                                               //Partner information is already known in the diagnostic structure
                                               IF (#diagnostics.partnerConfig.connnection.lifeSignCycleTime = T#0ms) THEN
                                                   //No --> Get diagnostics information
                                                   //LCom V2
                                                   IF (#statActualLocalLComVersion = #HEADER_V2) THEN
                                                       //UsesTimeStamp
                                                       #diagnostics.partnerConfig.timeSync.usePartnerTimestamps := BYTE_TO_BOOL(#statReceive.tempTelegram.data[2]);
                                                       //SendModeSyncTime
                                                       #diagnostics.partnerConfig.timeSync.sendMode := #statReceive.tempTelegram.data[3];
                                                       //LifeSignCycle
                                                       #tempDWord.%B3 := #statReceive.tempTelegram.data[4];
                                                       #tempDWord.%B2 := #statReceive.tempTelegram.data[5];
                                                       #tempDWord.%B1 := #statReceive.tempTelegram.data[6];
                                                       #tempDWord.%B0 := #statReceive.tempTelegram.data[7];
                                                       #statReceive.configTelegramV2.lifeSignCycle := DWORD_TO_TIME(#tempDWord);
                                                       #diagnostics.partnerConfig.connnection.lifeSignCycleTime := #statReceive.configTelegramV2.lifeSignCycle;
                                                       //Sender cycleTime
                                                       #tempDWord.%B3 := #statReceive.tempTelegram.data[8];
                                                       #tempDWord.%B2 := #statReceive.tempTelegram.data[9];
                                                       #tempDWord.%B1 := #statReceive.tempTelegram.data[10];
                                                       #tempDWord.%B0 := #statReceive.tempTelegram.data[11];
                                                       #statReceive.configTelegramV2.cycleTime := DWORD_TO_TIME(#tempDWord);
                                                       #diagnostics.partnerConfig.sender.cycleTime := #statReceive.configTelegramV2.cycleTime;
                                                       //Sender ackTimeOut
                                                       #tempDWord.%B3 := #statReceive.tempTelegram.data[12];
                                                       #tempDWord.%B2 := #statReceive.tempTelegram.data[13];
                                                       #tempDWord.%B1 := #statReceive.tempTelegram.data[14];
                                                       #tempDWord.%B0 := #statReceive.tempTelegram.data[15];
                                                       #statReceive.configTelegramV2.ackTimeOut := DWORD_TO_TIME(#tempDWord);
                                                       #diagnostics.partnerConfig.sender.ackTimeout := #statReceive.configTelegramV2.ackTimeOut;
                                                       //MaxSendDataLength
                                                       #tempDWord.%B3 := #statReceive.tempTelegram.data[16];
                                                       #tempDWord.%B2 := #statReceive.tempTelegram.data[17];
                                                       #tempDWord.%B1 := #statReceive.tempTelegram.data[18];
                                                       #tempDWord.%B0 := #statReceive.tempTelegram.data[19];
                                                       #statReceive.configTelegramV2.maxSendDataLength := #tempDWord;
                                                       #diagnostics.partnerConfig.sizeOfSendBuffer := #statReceive.configTelegramV2.maxSendDataLength;
                                                       //MaxReceiveDataLength
                                                       #tempDWord.%B3 := #statReceive.tempTelegram.data[20];
                                                       #tempDWord.%B2 := #statReceive.tempTelegram.data[21];
                                                       #tempDWord.%B1 := #statReceive.tempTelegram.data[22];
                                                       #tempDWord.%B0 := #statReceive.tempTelegram.data[23];
                                                       #statReceive.configTelegramV2.maxReceiveDataLength := #tempDWord;
                                                       #diagnostics.partnerConfig.sizeOfReceiveBuffer := #statReceive.configTelegramV2.maxReceiveDataLength;
                                                   ELSE
                                                       //LCom V1
                                                       //LifeSignCycle
                                                       #statReceive.configTelegramV1.lifeSignCycle.%B1 := #statReceive.tempTelegram.data[8];
                                                       #statReceive.configTelegramV1.lifeSignCycle.%B0 := #statReceive.tempTelegram.data[9];
                                                       #diagnostics.partnerConfig.connnection.lifeSignCycleTime := UINT_TO_TIME(#statReceive.configTelegramV1.lifeSignCycle);
                                                       //MaxSendDataLength
                                                       #statReceive.configTelegramV1.maxSendDataLength.%B1 := #statReceive.tempTelegram.data[12];
                                                       #statReceive.configTelegramV1.maxSendDataLength.%B0 := #statReceive.tempTelegram.data[13];
                                                       #diagnostics.partnerConfig.sizeOfSendBuffer := #statReceive.configTelegramV1.maxSendDataLength;
                                                       //MaxReceiveDataLength
                                                       #statReceive.configTelegramV1.maxReceiveDataLength.%B1 := #statReceive.tempTelegram.data[14];
                                                       #statReceive.configTelegramV1.maxReceiveDataLength.%B0 := #statReceive.tempTelegram.data[15];
                                                       #diagnostics.partnerConfig.sizeOfReceiveBuffer := #statReceive.configTelegramV1.maxReceiveDataLength;
                                                       //UsesTimeStamp
                                                       #diagnostics.partnerConfig.timeSync.usePartnerTimestamps := BYTE_TO_BOOL(#statReceive.tempTelegram.data[10]);
                                                       //SendModeSyncTime
                                                       #diagnostics.partnerConfig.timeSync.sendMode := #statReceive.tempTelegram.data[11];
                                                   END_IF;
                                               END_IF;

                                           1://Telegram type 1

                                               //Reset index, so a new temp. LCom header can be built
                                               #statReceive.tempTelegram.index := 0;
                                               #statReceive.numberOfLComHeader := #statReceive.numberOfLComHeader + 1;

                                               //LCom V1
                                               //LifeSignCycle
                                               #statReceive.configTelegramV1.lifeSignCycle.%B1 := #statReceive.tempTelegram.data[8];
                                               #statReceive.configTelegramV1.lifeSignCycle.%B0 := #statReceive.tempTelegram.data[9];
                                               #diagnostics.partnerConfig.connnection.lifeSignCycleTime := UINT_TO_TIME(#statReceive.configTelegramV1.lifeSignCycle);
                                               //Receiver cycleTime from receiver
                                               #statReceive.configTelegramV1.cycleTime.%B1 := #statReceive.tempTelegram.data[4];
                                               #statReceive.configTelegramV1.cycleTime.%B0 := #statReceive.tempTelegram.data[5];
                                               //Receiver ackTimeOut from receiver
                                               #statReceive.configTelegramV1.ackTimeOut.%B1 := #statReceive.tempTelegram.data[6];
                                               #statReceive.configTelegramV1.ackTimeOut.%B0 := #statReceive.tempTelegram.data[7];

                                               //Are receive cycle time and current sender cycle time and receive ackTimeOut and current sender ackTimeOut equal ?
                                               IF ((#statReceive.configTelegramV1.cycleTime = (TIME_TO_UINT(#diagnostics.localConfig.sender.cycleTime)))
                                                   AND
                                                   (#statReceive.configTelegramV1.ackTimeOut = (TIME_TO_UINT(#diagnostics.localConfig.sender.ackTimeout))))
                                               THEN
                                                   ;//Yes equal --> Set FB.#connected and diagnostics information
                                               ELSE
                                                   //Not equal --> Compare values and prioritize
                                                   //Compare cycle time
                                                   IF (#statReceive.configTelegramV1.cycleTime > (TIME_TO_UINT(#diagnostics.localConfig.sender.cycleTime))) THEN
                                                       #statSend.configTelegramV1.cycleTime := #statReceive.configTelegramV1.cycleTime;
                                                   ELSE
                                                       ;//Actual sender cycleTime is bigger than the received sender cycleTime
                                                   END_IF;

                                                   //Compare acknowledge timeout
                                                   IF (#statReceive.configTelegramV1.ackTimeOut > (TIME_TO_UINT(#diagnostics.localConfig.sender.ackTimeout))) THEN
                                                       #statSend.configTelegramV1.ackTimeOut := #statReceive.configTelegramV1.ackTimeOut;
                                                   ELSE
                                                       ;//Actual acknowledge timeout is bigger than the received sender acknowledge timeout
                                                   END_IF;

                                                   //Update diagnostics information
                                                   #diagnostics.localConfig.sender.cycleTime := UINT_TO_TIME(#statReceive.configTelegramV1.cycleTime);
                                                   #diagnostics.localConfig.sender.ackTimeout := UINT_TO_TIME(#statReceive.configTelegramV1.ackTimeOut);

                                                   //Send telegram 2
                                                   #statSend.tsendFct.data[#statSend.tsendFct.dataOffset] := #statSend.configTelegramV1.LComVersion;
                                                   #statSend.tsendFct.data[#statSend.tsendFct.dataOffset + 1] := 16#02;
                                                   #statSend.tsendFct.data[#statSend.tsendFct.dataOffset + 2] := #statSend.configTelegramV1.comMode;
                                                   #statSend.tsendFct.data[#statSend.tsendFct.dataOffset + 3] := #statSend.configTelegramV1.slidingWindow;
                                                   //Cycle time
                                                   #statSend.tsendFct.data[#statSend.tsendFct.dataOffset + 4] := #statSend.configTelegramV1.cycleTime.%B1;
                                                   #statSend.tsendFct.data[#statSend.tsendFct.dataOffset + 5] := #statSend.configTelegramV1.cycleTime.%B0;
                                                   //Acknowledge timeout
                                                   #statSend.tsendFct.data[#statSend.tsendFct.dataOffset + 6] := #statSend.configTelegramV1.ackTimeOut.%B1;
                                                   #statSend.tsendFct.data[#statSend.tsendFct.dataOffset + 7] := #statSend.configTelegramV1.ackTimeOut.%B0;
                                                   //LifeSignCycle
                                                   #statSend.tsendFct.data[#statSend.tsendFct.dataOffset + 8] := #statSend.configTelegramV1.lifeSignCycle.%B1;
                                                   #statSend.tsendFct.data[#statSend.tsendFct.dataOffset + 9] := #statSend.configTelegramV1.lifeSignCycle.%B0;
                                                   //Status
                                                   #statSend.tsendFct.data[#statSend.tsendFct.dataOffset + 10] := #statSend.configTelegramV1.status;
                                                   //SendModeSyncTime
                                                   #statSend.tsendFct.data[#statSend.tsendFct.dataOffset + 11] := #statSend.configTelegramV1.sendModeSyncTime;
                                                   //MaxSendDataLength
                                                   #statSend.tsendFct.data[#statSend.tsendFct.dataOffset + 12] := #statSend.configTelegramV1.maxSendDataLength.%B1;
                                                   #statSend.tsendFct.data[#statSend.tsendFct.dataOffset + 13] := #statSend.configTelegramV1.maxSendDataLength.%B0;
                                                   //MaxReceiveDataLength
                                                   #statSend.tsendFct.data[#statSend.tsendFct.dataOffset + 14] := #statSend.configTelegramV1.maxReceiveDataLength.%B1;
                                                   #statSend.tsendFct.data[#statSend.tsendFct.dataOffset + 15] := #statSend.configTelegramV1.maxReceiveDataLength.%B0;
                                                   //Calculate offset in the tcp send buffer
                                                   #statSend.tsendFct.dataOffset := #statSend.tsendFct.dataOffset + 16;
                                                   #statState.sender := #SEND_CONFIG;
                                               END_IF;

                                               //Set FB.#connected and #diagnostics information
                                               #connected := #statConnected := TRUE;
                                               #diagnostics.statistics.LComProtocolUsed := TRUE;
                                               #diagnostics.statistics.activeLComVersion := #HEADER_V1;
                                               //Write diagnostics
                                               #statDiag.bufferIndex := #statDiag.bufferIndex + 1;
                                               #statDiag.buffer[#statDiag.bufferIndex].status := #STATUS_CONNECTED_V1;
                                               #statDiag.buffer[#statDiag.bufferIndex].subFunctionErrorID := 16#0000;
                                               #statDiag.buffer[#statDiag.bufferIndex].additionalValue1 := 0.0;
                                               #statDiag.buffer[#statDiag.bufferIndex].additionalValue2 := 0.0;
                                               #statDiag.buffer[#statDiag.bufferIndex].additionalValue3 := 0.0;
                                               #statDiag.buffer[#statDiag.bufferIndex].additionalValue4 := T#0ms;

                                               #statState.cfgSender := #OPERATION;

                                               //MaxSendDataLength
                                               #statReceive.configTelegramV1.maxSendDataLength.%B1 := #statReceive.tempTelegram.data[12];
                                               #statReceive.configTelegramV1.maxSendDataLength.%B0 := #statReceive.tempTelegram.data[13];
                                               #diagnostics.partnerConfig.sizeOfSendBuffer := #statReceive.configTelegramV1.maxSendDataLength;
                                               //MaxReceiveDataLength
                                               #statReceive.configTelegramV1.maxReceiveDataLength.%B1 := #statReceive.tempTelegram.data[14];
                                               #statReceive.configTelegramV1.maxReceiveDataLength.%B0 := #statReceive.tempTelegram.data[15];
                                               #diagnostics.partnerConfig.sizeOfReceiveBuffer := #statReceive.configTelegramV1.maxReceiveDataLength;
                                               //UsesTimeStamp
                                               #diagnostics.partnerConfig.timeSync.usePartnerTimestamps := BYTE_TO_BOOL(#statReceive.tempTelegram.data[10]);
                                               //SendModeSyncTime
                                               #diagnostics.partnerConfig.timeSync.sendMode := #statReceive.tempTelegram.data[11];

                                               IF ((#diagnostics.localConfig.timeSync.usePartnerTimestamps
                                                   XOR
                                                   #diagnostics.partnerConfig.timeSync.usePartnerTimestamps)
                                                   AND
                                                   (#diagnostics.localConfig.timeSync.sendMode > 0
                                                   OR
                                                   #diagnostics.partnerConfig.timeSync.sendMode > 0))
                                               THEN
                                                   ;//One cpu does send timeSync information
                                               ELSE
                                                   //Write diagnostics
                                                   #statDiag.bufferIndex := #statDiag.bufferIndex + 1;
                                                   #statDiag.buffer[#statDiag.bufferIndex].status := #WARN_NO_TIME_SYNC;
                                                   #statDiag.buffer[#statDiag.bufferIndex].subFunctionErrorID := 16#0000;
                                                   #statDiag.buffer[#statDiag.bufferIndex].additionalValue1 := 0.0;
                                                   #statDiag.buffer[#statDiag.bufferIndex].additionalValue2 := 0.0;
                                                   #statDiag.buffer[#statDiag.bufferIndex].additionalValue3 := 0.0;
                                                   #statDiag.buffer[#statDiag.bufferIndex].additionalValue4 := T#0ms;
                                               END_IF;

                                           2://telegram type 2

                                               //Reset index, so a new temp. LCom header can be built
                                               #statReceive.tempTelegram.index := 0;
                                               #statReceive.numberOfLComHeader := #statReceive.numberOfLComHeader + 1;

                                               //LCom V2
                                               IF (#statActualLocalLComVersion = #HEADER_V2) THEN
                                                   //UsesTimeStamp
                                                   #diagnostics.partnerConfig.timeSync.usePartnerTimestamps := BYTE_TO_BOOL(#statReceive.tempTelegram.data[2]);
                                                   //SendModeSyncTime
                                                   #diagnostics.partnerConfig.timeSync.sendMode := #statReceive.tempTelegram.data[3];
                                                   //LifeSignCycle
                                                   #tempDWord.%B3 := #statReceive.tempTelegram.data[4];
                                                   #tempDWord.%B2 := #statReceive.tempTelegram.data[5];
                                                   #tempDWord.%B1 := #statReceive.tempTelegram.data[6];
                                                   #tempDWord.%B0 := #statReceive.tempTelegram.data[7];
                                                   #statReceive.configTelegramV2.lifeSignCycle := DWORD_TO_TIME(#tempDWord);
                                                   #diagnostics.partnerConfig.connnection.lifeSignCycleTime := #statReceive.configTelegramV2.lifeSignCycle;

                                                   //Sender cycleTime
                                                   #tempDWord.%B3 := #statReceive.tempTelegram.data[8];
                                                   #tempDWord.%B2 := #statReceive.tempTelegram.data[9];
                                                   #tempDWord.%B1 := #statReceive.tempTelegram.data[10];
                                                   #tempDWord.%B0 := #statReceive.tempTelegram.data[11];
                                                   #statReceive.configTelegramV2.cycleTime := DWORD_TO_TIME(#tempDWord);
                                                   #diagnostics.partnerConfig.sender.cycleTime := #statReceive.configTelegramV2.cycleTime;
                                                   //Sender ackTimeOut
                                                   #tempDWord.%B3 := #statReceive.tempTelegram.data[12];
                                                   #tempDWord.%B2 := #statReceive.tempTelegram.data[13];
                                                   #tempDWord.%B1 := #statReceive.tempTelegram.data[14];
                                                   #tempDWord.%B0 := #statReceive.tempTelegram.data[15];
                                                   #statReceive.configTelegramV2.ackTimeOut := DWORD_TO_TIME(#tempDWord);
                                                   #diagnostics.partnerConfig.sender.ackTimeout := #statReceive.configTelegramV2.ackTimeOut;
                                                   //MaxSendDataLength
                                                   #tempDWord.%B3 := #statReceive.tempTelegram.data[16];
                                                   #tempDWord.%B2 := #statReceive.tempTelegram.data[17];
                                                   #tempDWord.%B1 := #statReceive.tempTelegram.data[18];
                                                   #tempDWord.%B0 := #statReceive.tempTelegram.data[19];
                                                   #statReceive.configTelegramV2.maxSendDataLength := #tempDWord;
                                                   #diagnostics.partnerConfig.sizeOfSendBuffer := #statReceive.configTelegramV2.maxSendDataLength;
                                                   //MaxReceiveDataLength
                                                   #tempDWord.%B3 := #statReceive.tempTelegram.data[20];
                                                   #tempDWord.%B2 := #statReceive.tempTelegram.data[21];
                                                   #tempDWord.%B1 := #statReceive.tempTelegram.data[22];
                                                   #tempDWord.%B0 := #statReceive.tempTelegram.data[23];
                                                   #statReceive.configTelegramV2.maxReceiveDataLength := #tempDWord;
                                                   #diagnostics.partnerConfig.sizeOfReceiveBuffer := #statReceive.configTelegramV2.maxReceiveDataLength;

                                                   //Set FB.#connected and #diagnostics information
                                                   #connected := #statConnected := TRUE;
                                                   #diagnostics.statistics.LComProtocolUsed := TRUE;
                                                   #diagnostics.statistics.activeLComVersion := #HEADER_V2;
                                                   #statState.cfgSender := #OPERATION;

                                                   //Write diagnostics
                                                   #statDiag.bufferIndex := #statDiag.bufferIndex + 1;
                                                   #statDiag.buffer[#statDiag.bufferIndex].status := #STATUS_CONNECTED_V2;
                                                   #statDiag.buffer[#statDiag.bufferIndex].subFunctionErrorID := 16#0000;
                                                   #statDiag.buffer[#statDiag.bufferIndex].additionalValue1 := 0.0;
                                                   #statDiag.buffer[#statDiag.bufferIndex].additionalValue2 := 0.0;
                                                   #statDiag.buffer[#statDiag.bufferIndex].additionalValue3 := 0.0;
                                                   #statDiag.buffer[#statDiag.bufferIndex].additionalValue4 := T#0ms;

                                                   //Check timeSync setting at local cpu and partner cpu
                                                   IF ((#diagnostics.localConfig.timeSync.usePartnerTimestamps
                                                       XOR
                                                       #diagnostics.partnerConfig.timeSync.usePartnerTimestamps)
                                                       AND
                                                       (#diagnostics.localConfig.timeSync.sendMode > 0
                                                       OR
                                                       #diagnostics.partnerConfig.timeSync.sendMode > 0))
                                                   THEN
                                                       ;//One cpu does send timeSync information
                                                   ELSE
                                                       //Write diagnostics
                                                       #statDiag.bufferIndex := #statDiag.bufferIndex + 1;
                                                       #statDiag.buffer[#statDiag.bufferIndex].status := #WARN_NO_TIME_SYNC;
                                                       #statDiag.buffer[#statDiag.bufferIndex].subFunctionErrorID := 16#0000;
                                                       #statDiag.buffer[#statDiag.bufferIndex].additionalValue1 := 0.0;
                                                       #statDiag.buffer[#statDiag.bufferIndex].additionalValue2 := 0.0;
                                                       #statDiag.buffer[#statDiag.bufferIndex].additionalValue3 := 0.0;
                                                       #statDiag.buffer[#statDiag.bufferIndex].additionalValue4 := T#0ms;
                                                   END_IF;
                                                   //Do not send telegram 1
                                               ELSE
                                                   //LCom V1
                                                   //LifeSignCycle
                                                   #statReceive.configTelegramV1.lifeSignCycle.%B1 := #statReceive.tempTelegram.data[8];
                                                   #statReceive.configTelegramV1.lifeSignCycle.%B0 := #statReceive.tempTelegram.data[9];
                                                   #diagnostics.partnerConfig.connnection.lifeSignCycleTime := UINT_TO_TIME(#statReceive.configTelegramV1.lifeSignCycle);
                                                   //CycleTime
                                                   #statReceive.configTelegramV1.cycleTime.%B1 := #statReceive.tempTelegram.data[4];
                                                   #statReceive.configTelegramV1.cycleTime.%B0 := #statReceive.tempTelegram.data[5];
                                                   #diagnostics.partnerConfig.sender.cycleTime := UINT_TO_TIME(#statReceive.configTelegramV1.cycleTime);
                                                   //AckTimeOut
                                                   #statReceive.configTelegramV1.ackTimeOut.%B1 := #statReceive.tempTelegram.data[6];
                                                   #statReceive.configTelegramV1.ackTimeOut.%B0 := #statReceive.tempTelegram.data[7];
                                                   #diagnostics.partnerConfig.sender.ackTimeout := UINT_TO_TIME(#statReceive.configTelegramV1.ackTimeOut);
                                                   //MaxSendDataLength
                                                   #statReceive.configTelegramV1.maxSendDataLength.%B1 := #statReceive.tempTelegram.data[12];
                                                   #statReceive.configTelegramV1.maxSendDataLength.%B0 := #statReceive.tempTelegram.data[13];
                                                   #diagnostics.partnerConfig.sizeOfSendBuffer := #statReceive.configTelegramV1.maxSendDataLength;
                                                   //MaxReceiveDataLength
                                                   #statReceive.configTelegramV1.maxReceiveDataLength.%B1 := #statReceive.tempTelegram.data[14];
                                                   #statReceive.configTelegramV1.maxReceiveDataLength.%B0 := #statReceive.tempTelegram.data[15];
                                                   #diagnostics.partnerConfig.sizeOfReceiveBuffer := #statReceive.configTelegramV1.maxReceiveDataLength;
                                                   //UsesTimeStamp
                                                   #diagnostics.partnerConfig.timeSync.usePartnerTimestamps := BYTE_TO_BOOL(#statReceive.tempTelegram.data[10]);
                                                   //SendModeSyncTime
                                                   #diagnostics.partnerConfig.timeSync.sendMode := #statReceive.tempTelegram.data[11];

                                                   //Send Telegram 1
                                                   #statSend.tsendFct.data[#statSend.tsendFct.dataOffset] := #statSend.configTelegramV1.LComVersion;
                                                   #statSend.tsendFct.data[#statSend.tsendFct.dataOffset + 1] := 16#01;
                                                   #statSend.tsendFct.data[#statSend.tsendFct.dataOffset + 2] := #statSend.configTelegramV1.comMode;
                                                   #statSend.tsendFct.data[#statSend.tsendFct.dataOffset + 3] := #statSend.configTelegramV1.slidingWindow;
                                                   //CycleTime
                                                   #statSend.tsendFct.data[#statSend.tsendFct.dataOffset + 4] := #statReceive.configTelegramV1.cycleTime.%B1;
                                                   #statSend.tsendFct.data[#statSend.tsendFct.dataOffset + 5] := #statReceive.configTelegramV1.cycleTime.%B0;
                                                   //AckTimeOut
                                                   #statSend.tsendFct.data[#statSend.tsendFct.dataOffset + 6] := #statReceive.configTelegramV1.ackTimeOut.%B1;
                                                   #statSend.tsendFct.data[#statSend.tsendFct.dataOffset + 7] := #statReceive.configTelegramV1.ackTimeOut.%B0;
                                                   //LifeSignCycle
                                                   #statSend.tsendFct.data[#statSend.tsendFct.dataOffset + 8] := #statSend.configTelegramV1.lifeSignCycle.%B1;
                                                   #statSend.tsendFct.data[#statSend.tsendFct.dataOffset + 9] := #statSend.configTelegramV1.lifeSignCycle.%B0;
                                                   //Status
                                                   #statSend.tsendFct.data[#statSend.tsendFct.dataOffset + 10] := #statSend.configTelegramV1.status;
                                                   //SendModeSyncTime
                                                   #statSend.tsendFct.data[#statSend.tsendFct.dataOffset + 11] := #statSend.configTelegramV1.sendModeSyncTime;
                                                   //MaxSendDataLength
                                                   #statSend.tsendFct.data[#statSend.tsendFct.dataOffset + 12] := #statSend.configTelegramV1.maxSendDataLength.%B1;
                                                   #statSend.tsendFct.data[#statSend.tsendFct.dataOffset + 13] := #statSend.configTelegramV1.maxSendDataLength.%B0;
                                                   //MaxReceiveDataLength
                                                   #statSend.tsendFct.data[#statSend.tsendFct.dataOffset + 14] := #statSend.configTelegramV1.maxReceiveDataLength.%B1;
                                                   #statSend.tsendFct.data[#statSend.tsendFct.dataOffset + 15] := #statSend.configTelegramV1.maxReceiveDataLength.%B0;
                                                   //Calculate offset in the tcp send buffer
                                                   #statSend.tsendFct.dataOffset := #statSend.tsendFct.dataOffset + 16;
                                                   //Set state
                                                   #statState.sender := #SEND_CONFIG;
                                               END_IF;

                                           5://Telegram type 5

                                               //Reset index, so a new temp. LCom header can be built
                                               #statReceive.tempTelegram.index := 0;
                                               #statReceive.numberOfLComHeader := #statReceive.numberOfLComHeader + 1;

                                               //Accept timestamp from partner ?
                                               IF (#diagnostics.localConfig.timeSync.usePartnerTimestamps) THEN
                                                   //Yes --> Accept timestamp from partner
                                                   #tempActTime.YEAR := INT_TO_UINT(BCD16_TO_INT(#statReceive.tempTelegram.data[2] AND 16#00FF));
                                                   IF ((#tempActTime.YEAR >= 90)
                                                       AND (#tempActTime.YEAR <= 99))
                                                   THEN
                                                       #tempActTime.YEAR := #tempActTime.YEAR + 1900;
                                                   ELSE
                                                       #tempActTime.YEAR := #tempActTime.YEAR + 2000;
                                                   END_IF;

                                                   #tempActTime.MONTH := INT_TO_USINT(BCD16_TO_INT(#statReceive.tempTelegram.data[3] AND 16#00FF));
                                                   #tempActTime.DAY := INT_TO_USINT(BCD16_TO_INT(#statReceive.tempTelegram.data[4] AND 16#00FF));
                                                   #tempActTime.HOUR := INT_TO_USINT(BCD16_TO_INT(#statReceive.tempTelegram.data[5] AND 16#00FF));
                                                   #tempActTime.MINUTE := INT_TO_USINT(BCD16_TO_INT(#statReceive.tempTelegram.data[6] AND 16#00FF));
                                                   #tempActTime.SECOND := INT_TO_USINT(BCD16_TO_INT(#statReceive.tempTelegram.data[7] AND 16#00FF));
                                                   #tempActTime.NANOSECOND := INT_TO_UDINT(BCD16_TO_INT(#statReceive.tempTelegram.data[8] AND 16#00FF));
                                                   #tempActTime.NANOSECOND := #tempActTime.NANOSECOND * 1000;
                                                   #tempActTime.NANOSECOND := #tempActTime.NANOSECOND + 500;
                                                   #tempActTime.WEEKDAY := INT_TO_USINT(BCD16_TO_INT(#statReceive.tempTelegram.data[9] AND 16#000F));
                                                   //Write local time
                                                   #statRet := WR_LOC_T(LOCTIME := #tempActTime, DST := FALSE);
                                                   //Statistic --> Get time stamp of last time sync
                                                   #diagnostics.statistics.lastTimeSync := #tempActTime;
                                               ELSE
                                                   ;//No --> Do not write system time
                                               END_IF;

                                           20://Telegram type 20

                                               //Reset index, so a new temp. LCom header can be built
                                               #statReceive.numberOfLComHeader := #statReceive.numberOfLComHeader + 1;
                                               #statReceive.tempTelegram.index := 0;

                                               //Write diagnostics ---> Stop analyzing the tcp receive buffer
                                               #statDiag.bufferIndex := #statDiag.bufferIndex + 1;
                                               #statDiag.buffer[#statDiag.bufferIndex].status := #STATUS_DISCONNECTING;
                                               #statDiag.buffer[#statDiag.bufferIndex].subFunctionErrorID := 16#0000;
                                               #statDiag.buffer[#statDiag.bufferIndex].additionalValue1 := 0.0;
                                               #statDiag.buffer[#statDiag.bufferIndex].additionalValue2 := 0.0;
                                               #statDiag.buffer[#statDiag.bufferIndex].additionalValue3 := 0.0;
                                               #statDiag.buffer[#statDiag.bufferIndex].additionalValue4 := T#0ms;
                                               #statState.connection := #CLOSE_CONNECTION;
                                               EXIT;

                                           ELSE//Telegram type is unknown
                                               //Write diagnostics
                                               #statDiag.bufferIndex := #statDiag.bufferIndex + 1;
                                               #statDiag.buffer[#statDiag.bufferIndex].status := #ERR_WRONG_TELEGRAM_ID;
                                               #statDiag.buffer[#statDiag.bufferIndex].subFunctionErrorID := 16#0000;
                                               #statDiag.buffer[#statDiag.bufferIndex].additionalValue1 := #statReceive.tempTelegram.telegramType;
                                               #statDiag.buffer[#statDiag.bufferIndex].additionalValue2 := 0.0;
                                               #statDiag.buffer[#statDiag.bufferIndex].additionalValue3 := 0.0;
                                               #statDiag.buffer[#statDiag.bufferIndex].additionalValue4 := T#0ms;
                                               #statState.connection := #CLOSE_CONNECTION;
                                               GOTO diag;
                                       END_CASE;

                                   END_IF;
                               END_REGION LCOM_PROTOCOL

                               //Calculate rest of data in the tcp receive buffer
                               #statReceive.trcvFct.dataLengthRest := #statReceive.trcvFct.dataLength - #statReceive.trcvFct.dataOffset;

                           UNTIL ((#statReceive.trcvFct.dataLengthRest <= 0)
                               OR (#statReceive.trcvFct.dataLengthRest > #MAX_DATA_BUFFER))
                               //If the result of the calculation of the rest data is greater than 4096, then an error occurred
                           END_REPEAT;
                           //End:Analyze tcp receive buffer with LCom protocol

                       END_IF;//#readDataLength <> 0
                   END_REGION READ_TCP_BUFFER

                   REGION HANDLE_SENDING
                       //---------------------------------------------------------------------
                       //Check if next package can be sent
                       //---------------------------------------------------------------------
                       IF ((#statConnected = TRUE) AND (#statState.connection = #OPERATION)) THEN

                           //Get cycle time [ms]
                           #instLocalCycleTimeTimer(IN := TRUE,
                                                    PT := #diagnostics.localConfig.sender.cycleTime);


                           //---------------------------------------------------------------------
                           //In sending process
                           //---------------------------------------------------------------------
                           IF (#statSending = TRUE) THEN
                               //Yes --> In sending process

                               REGION CHECK_SEND_CYCLETIME
                                   //---------------------------------------------------------------------
                                   //Check if sender cycle time is expired (with and without LCom protocol) ?
                                   //---------------------------------------------------------------------
                                   IF (#instLocalCycleTimeTimer.Q AND #diagnostics.localConfig.sender.cycleTime > T#0ms) THEN
                                       //Yes --> Sender cycle time is expired
                                       //Check if sender cycle time violation is already stored ?
                                       IF (#statSend.userData.sendCycleViolation) THEN
                                           ;//Yes --> Exceeded before and stored
                                       ELSE
                                           //No --> Increase number of send cycle time violations
                                           #diagnostics.statistics.totalSendCycleViolations := #diagnostics.statistics.totalSendCycleViolations + 1;
                                           #statSend.userData.sendCycleViolation := TRUE;
                                       END_IF;

                                       //Write diagnostics
                                       #statDiag.bufferIndex := #statDiag.bufferIndex + 1;
                                       #statDiag.buffer[#statDiag.bufferIndex].status := #WARN_SEND_CYCLE_EXPIRED;
                                       #statDiag.buffer[#statDiag.bufferIndex].subFunctionErrorID := 16#0000;
                                       #statDiag.buffer[#statDiag.bufferIndex].additionalValue1 := UDINT_TO_REAL(TIME_TO_UDINT(#diagnostics.localConfig.sender.cycleTime));
                                       #statDiag.buffer[#statDiag.bufferIndex].additionalValue2 := 0.0;
                                       #statDiag.buffer[#statDiag.bufferIndex].additionalValue3 := 0.0;
                                       #statDiag.buffer[#statDiag.bufferIndex].additionalValue4 := #instLocalCycleTimeTimer.ET;
                                   ELSE
                                       ;//No --> Sender cycle time is not expired
                                   END_IF;//End: Check if sender cycle time is expired (with and without LCom protocol) ?
                               END_REGION CHECK_SEND_CYCLETIME

                               REGION CHECK_ACK_TIMEOUT
                                   //---------------------------------------------------------------------
                                   //Check acknowledge timeout with LCom protocol
                                   //---------------------------------------------------------------------
                                   IF (#diagnostics.localConfig.connection.useLComProtocol = TRUE) THEN

                                       //Get acknowledge timeout [ms]
                                       #instExpectedAckPackage1(IN := TRUE,
                                                                PT := #diagnostics.localConfig.sender.ackTimeout);

                                       //Check if acknowledge timeout is expired ?
                                       IF ((#instExpectedAckPackage1.Q = TRUE)
                                           AND
                                           (#statSend.numberOfLComPackage > 0))
                                       THEN
                                           //Yes --> Acknowledge timeout is expired, increase number of confirmation timeouts
                                           #diagnostics.statistics.totalAckTimeouts := #diagnostics.statistics.totalAckTimeouts + 1;

                                           //Write diagnostics
                                           #statDiag.bufferIndex := #statDiag.bufferIndex + 1;
                                           #statDiag.buffer[#statDiag.bufferIndex].status := #ERR_ACK_TIMEOUT_EXPIRED;
                                           #statDiag.buffer[#statDiag.bufferIndex].subFunctionErrorID := 16#0000;
                                           #statDiag.buffer[#statDiag.bufferIndex].additionalValue1 := UDINT_TO_REAL(TIME_TO_UDINT(#diagnostics.localConfig.sender.ackTimeout));
                                           #statDiag.buffer[#statDiag.bufferIndex].additionalValue2 := 0.0;
                                           #statDiag.buffer[#statDiag.bufferIndex].additionalValue3 := 0.0;
                                           #statDiag.buffer[#statDiag.bufferIndex].additionalValue4 := #instExpectedAckPackage1.ET;
                                           #statState.connection := #CLOSE_CONNECTION;
                                           GOTO diag;
                                       ELSE
                                           //No --> Acknowledge timeout is not expired

                                           //Is the last LCom package already sent ?
                                           IF (#statState.comSender = #SEND_NO_DATA) THEN
                                               ;//Yes --> Wait for acknowledge telegram
                                           ELSE
                                               //No --> Last LCom package not sent yet

                                               //Check if the next LCom package can be sent ? (Sliding window)
                                               IF ((#statSend.numberOfLComPackage < 1)
                                                   AND
                                                   (#diagnostics.statistics.activeLComVersion = #HEADER_V1
                                                   OR
                                                   #diagnostics.statistics.activeLComVersion = #HEADER_V2))
                                               THEN
                                                   //Yes --> Continue sending
                                                   #statState.comSender := #CYCLE;
                                               ELSE
                                                   //No --> Wait for acknowledge telegram
                                                   #statState.comSender := #WAIT_ACK_TELEGRAM;
                                               END_IF;
                                           END_IF;//End: Is the last LCom package already sent ?
                                       END_IF;//End: Check if acknowledge time is expired ?
                                   ELSE
                                       //Continue without LCom protocol, acknowledge timeout is not valid
                                       #statState.comSender := #CYCLE;
                                   END_IF;
                               END_REGION CHECK_ACK_TIMEOUT

                           ELSE
                               //Not --> Not in sending process
                               REGION CHECK_SEND_CONFIG_AND_DATA_TO_SEND
                                   //With LCom protocol --> Check if sender configuration was changed
                                   IF (#diagnostics.localConfig.connection.useLComProtocol = TRUE
                                       AND
                                       ((#configuration.sender.cycleTime <> #statCompare.sender.cycleTime)
                                       OR
                                       (#configuration.sender.ackTimeout <> #statCompare.sender.ackTimeOut)))
                                   THEN
                                       #connected := #statConnected := FALSE;
                                       //Update parameters
                                       #statState.cfgSender := #STATE_INIT;
                                   ELSIF (NOT #diagnostics.localConfig.connection.useLComProtocol
                                       AND
                                       #configuration.sender.cycleTime <> #statCompare.sender.cycleTime)
                                   THEN//Without LCom protocol --> Check if sender configuration was changed
                                       //Update parameters
                                       #diagnostics.localConfig.sender.cycleTime := #configuration.sender.cycleTime;
                                       #statCompare.sender.cycleTime := #configuration.sender.cycleTime;
                                   ELSIF (#send OR #statRisingEdgeSend)//Check if FB.send input is true or rising edge is detected ?
                                   THEN
                                       //Yes --> FB.send input is true

                                       //---------------------------------------------------------------------
                                       //Check if data have to be sent
                                       //---------------------------------------------------------------------
                                       IF ((#sendDataLength > 0)
                                           AND
                                           ((#statRisingEdgeSend)//Rising edge
                                           OR
                                           ((#instLocalCycleTimeTimer.Q)//check CycleTimeTimer
                                           AND
                                           (#diagnostics.localConfig.sender.cycleTime > T#0ms))))
                                       THEN
                                           //Start sending
                                           #sending := #statSending := TRUE;
                                           #statSend.userData.sendCycleViolation := FALSE;
                                           #statSend.userData.offset := 0;
                                           #statRisingEdgeSend := FALSE;

                                           //Start message sending timer
                                           #instMsgSendingTimer(IN := TRUE,
                                                                PT := T#+24d20h31m23s647ms);

                                           //Stop/Start local cycle timer
                                           #instLocalCycleTimeTimer(IN := FALSE,
                                                                    PT := #diagnostics.localConfig.sender.cycleTime);
                                           #instLocalCycleTimeTimer(IN := TRUE,
                                                                    PT := #diagnostics.localConfig.sender.cycleTime);


                                           //Send data length greater than size of local send buffer ?
                                           IF (#sendDataLength > #diagnostics.localConfig.sizeOfSendBuffer) THEN
                                               //Yes --> Send data length is greater than size of local send buffer
                                               #statSend.dataTelegram.totalMessageLength := #diagnostics.localConfig.sizeOfSendBuffer;

                                               IF #diagnostics.localConfig.connection.useLComProtocol THEN
                                                   #statSend.dataTelegram.totalMessageLength := #diagnostics.localConfig.sizeOfSendBuffer;
                                               ELSE
                                                   #statSend.dataTelegram.totalMessageLength := #sendDataLength;
                                               END_IF;
                                               //Write diagnostics
                                               #statDiag.bufferIndex := #statDiag.bufferIndex + 1;
                                               #statDiag.buffer[#statDiag.bufferIndex].status := #WARN_SEND_DATA_LENGTH;
                                               #statDiag.buffer[#statDiag.bufferIndex].subFunctionErrorID := 16#0000;
                                               #statDiag.buffer[#statDiag.bufferIndex].additionalValue1 := UDINT_TO_REAL(#sendDataLength);
                                               #statDiag.buffer[#statDiag.bufferIndex].additionalValue2 := UDINT_TO_REAL(#diagnostics.localConfig.sizeOfSendBuffer);
                                               #statDiag.buffer[#statDiag.bufferIndex].additionalValue3 := 0.0;
                                               #statDiag.buffer[#statDiag.bufferIndex].additionalValue4 := T#0ms;
                                           ELSE
                                               //No --> Send data length is less than size of local send buffer
                                               #statSend.dataTelegram.totalMessageLength := #sendDataLength;
                                           END_IF;

                                           //"Send data length" greater than size of partner receive buffer ?
                                           IF ((#diagnostics.localConfig.connection.useLComProtocol)
                                               AND
                                               (#diagnostics.partnerConfig.sizeOfReceiveBuffer < #statSend.dataTelegram.totalMessageLength)
                                               ) THEN
                                               //Yes --> "Send data length" is greater than size of partner receive buffer
                                               #statSend.dataTelegram.totalMessageLength := #diagnostics.partnerConfig.sizeOfReceiveBuffer;
                                               //Write diagnostics
                                               #statDiag.bufferIndex := #statDiag.bufferIndex + 1;
                                               #statDiag.buffer[#statDiag.bufferIndex].status := #WARN_RECEIVE_BUFFER_LEN;
                                               #statDiag.buffer[#statDiag.bufferIndex].subFunctionErrorID := 16#0000;
                                               #statDiag.buffer[#statDiag.bufferIndex].additionalValue1 := UDINT_TO_REAL(#sendDataLength);
                                               #statDiag.buffer[#statDiag.bufferIndex].additionalValue2 := UDINT_TO_REAL(#diagnostics.partnerConfig.sizeOfReceiveBuffer);
                                               #statDiag.buffer[#statDiag.bufferIndex].additionalValue3 := 0.0;
                                               #statDiag.buffer[#statDiag.bufferIndex].additionalValue4 := T#0ms;
                                           ELSE
                                               ;//No --> "Send data length" is less than size of partner receive buffer
                                           END_IF;

                                           //Increase message counter
                                           #statSend.dataTelegram.messageCounter := #statSend.dataTelegram.messageCounter + 1;

                                           #statState.comSender := #CYCLE;
                                       ELSE
                                           //Cycle time is not expired
                                           #statState.comSender := #STATE_WAIT;
                                       END_IF;//End: Check if data have to be send ?
                                   ELSE
                                       //Sender configuration was not changed
                                       //FB:send = FALSE
                                       #statState.comSender := #STATE_INACTIVE;
                                       #statOldSend := FALSE;
                                   END_IF;
                               END_REGION CHECK_SEND_CONFIG_AND_DATA_TO_SEND

                               //Update
                               #statCompare.sender.cycleTime := #configuration.sender.cycleTime;
                               #statCompare.sender.ackTimeOut := #configuration.sender.ackTimeout;

                               REGION TIME_SYNCHRONIZATION
                                   //---------------------------------------------------------------------
                                   //Time synchronization
                                   //---------------------------------------------------------------------

                                   //Calculate rest bytes from tcp send buffer
                                   #statSend.tsendFct.dataLengthRest := (#MAX_DATA_BUFFER - #statSend.tsendFct.dataOffset);

                                   //---------------------------------------------------------------------
                                   //10 Bytes still free in the tcp send buffer
                                   //---------------------------------------------------------------------
                                   IF ((#diagnostics.localConfig.connection.useLComProtocol)
                                       AND
                                       (#diagnostics.localConfig.timeSync.sendMode > 0)
                                       AND
                                       (NOT (#diagnostics.localConfig.timeSync.usePartnerTimestamps))
                                       AND
                                       (#diagnostics.partnerConfig.timeSync.usePartnerTimestamps)
                                       AND
                                       (#statSend.tsendFct.dataLengthRest >= 10))
                                   THEN
                                       //Yes 10 bytes still free --> Get local time
                                       #statRet := RD_LOC_T(#tempActTime);

                                       CASE #diagnostics.localConfig.timeSync.sendMode OF
                                           0:
                                               ;//Time synchronization is inactive

                                           1: //Cycle time synchronization --> Get cycle time [ms]

                                               #instSyncTimer(IN := TRUE,
                                                              PT := #diagnostics.localConfig.timeSync.cycleTime);

                                               //Cycle time expired ?
                                               IF ((#instSyncTimer.Q) OR (#diagnostics.statistics.lastTimeSync.YEAR = 2200)) THEN
                                                   //Stop/Start local cycle timer
                                                   #instSyncTimer(IN := FALSE,
                                                                  PT := #diagnostics.localConfig.timeSync.cycleTime);
                                                   #instSyncTimer(IN := TRUE,
                                                                  PT := #diagnostics.localConfig.timeSync.cycleTime);
                                                   //Statistic --> Get time stamp of last time sync
                                                   #diagnostics.statistics.lastTimeSync := #tempActTime;
                                               END_IF;
                                           2: //Time of day synchronization
                                               IF ((DTL_TO_TOD(#tempActTime) > #diagnostics.localConfig.timeSync.sendAtTimeOfDay)
                                                   OR
                                                   #diagnostics.statistics.lastTimeSync.YEAR = 2200)
                                               THEN

                                                   IF #diagnostics.statistics.lastTimeSync.YEAR = 2200 THEN
                                                       //Start after connect
                                                       #diagnostics.statistics.lastTimeSync := #tempActTime;
                                                       //Is the date unequal
                                                   ELSIF (#diagnostics.statistics.lastTimeSync.DAY <> #tempActTime.DAY) THEN
                                                       //Yes --> date is unequal
                                                       #diagnostics.statistics.lastTimeSync := #tempActTime;
                                                   ELSE
                                                       //No --> date is equal
                                                       //Has the time sync telegram already sent on specified time of day ?
                                                       IF (DTL_TO_TOD(#diagnostics.statistics.lastTimeSync) > #diagnostics.localConfig.timeSync.sendAtTimeOfDay) THEN
                                                           ;//already sent, nothing to do
                                                       ELSE
                                                           #diagnostics.statistics.lastTimeSync := #tempActTime;
                                                       END_IF;
                                                   END_IF;
                                               END_IF;
                                           ELSE
                                               ;
                                       END_CASE;

                                       //Build telegram 5 (time synchronization) ?
                                       IF (#diagnostics.statistics.lastTimeSync = #tempActTime) THEN

                                           #statSend.tsendFct.data[#statSend.tsendFct.dataOffset] := #diagnostics.statistics.activeLComVersion;
                                           #statSend.tsendFct.data[#statSend.tsendFct.dataOffset + 1] := 16#05;

                                           //Convert from nSecond in mSecond
                                           #tempActTime.NANOSECOND := #tempActTime.NANOSECOND / 1000000;
                                           #statSend.tsendFct.data[#statSend.tsendFct.dataOffset + 8] := WORD_TO_BYTE(SHR(N := 4, IN := ((INT_TO_BCD16(UDINT_TO_INT(#tempActTime.NANOSECOND))))));

                                           #statSend.tsendFct.data[#statSend.tsendFct.dataOffset + 3] := WORD_TO_BYTE(INT_TO_BCD16(UDINT_TO_INT(#tempActTime.NANOSECOND)) AND 16#000F);
                                           #statSend.tsendFct.data[#statSend.tsendFct.dataOffset + 9] := SHL(IN := #statSend.tsendFct.data[#statSend.tsendFct.dataOffset + 3], N := 4);
                                           #statSend.tsendFct.data[#statSend.tsendFct.dataOffset + 2] := WORD_TO_BYTE(INT_TO_BCD16(#tempActTime.WEEKDAY));
                                           #statSend.tsendFct.data[#statSend.tsendFct.dataOffset + 9] := #statSend.tsendFct.data[#statSend.tsendFct.dataOffset + 9] + #statSend.tsendFct.data[#statSend.tsendFct.dataOffset + 2];


                                           IF ((#tempActTime.YEAR > 1970) AND (#tempActTime.YEAR <= 1990)) THEN
                                               #tempActTime.YEAR := 1990;
                                           ELSIF ((#tempActTime.YEAR > 1990) AND (#tempActTime.YEAR <= 1999)) THEN
                                               #tempActTime.YEAR := #tempActTime.YEAR - 1900;
                                           ELSE
                                               #tempActTime.YEAR := #tempActTime.YEAR - 2000;
                                           END_IF;

                                           #statSend.tsendFct.data[#statSend.tsendFct.dataOffset + 2] := WORD_TO_BYTE(INT_TO_BCD16(UINT_TO_INT(#tempActTime.YEAR)));
                                           #statSend.tsendFct.data[#statSend.tsendFct.dataOffset + 3] := WORD_TO_BYTE(INT_TO_BCD16(#tempActTime.MONTH));
                                           #statSend.tsendFct.data[#statSend.tsendFct.dataOffset + 4] := WORD_TO_BYTE(INT_TO_BCD16(#tempActTime.DAY));
                                           #statSend.tsendFct.data[#statSend.tsendFct.dataOffset + 5] := WORD_TO_BYTE(INT_TO_BCD16(#tempActTime.HOUR));
                                           #statSend.tsendFct.data[#statSend.tsendFct.dataOffset + 6] := WORD_TO_BYTE(INT_TO_BCD16(#tempActTime.MINUTE));
                                           #statSend.tsendFct.data[#statSend.tsendFct.dataOffset + 7] := WORD_TO_BYTE(INT_TO_BCD16(#tempActTime.SECOND));

                                           #statState.sender := #SEND_DATA;
                                           //Calculate offset in the tcp send buffer
                                           #statSend.tsendFct.dataOffset := #statSend.tsendFct.dataOffset + 10;
                                       END_IF;
                                   ELSE
                                       ;//No space
                                   END_IF;//End: 10 bytes still free in the tcp send buffer
                               END_REGION TIME_SYNCHRONIZATION

                           END_IF;//End: In sending process

                           REGION SEND_DATA_TELEGRAM
                               //---------------------------------------------------------------------
                               //Send telegram
                               //---------------------------------------------------------------------
                               IF (#statState.comSender = #CYCLE
                                   AND
                                   (#diagnostics.localConfig.connection.useLComProtocol))
                               THEN
                                   //---------------------------------------------------------------------
                                   //Send data telegram with LCom protocol
                                   //---------------------------------------------------------------------
                                   #statState.sender := #SEND_DATA;

                                   //Calculate rest bytes from tcp send buffer
                                   IF (#diagnostics.statistics.activeLComVersion = #HEADER_V2) THEN
                                       #statSend.tsendFct.dataLengthRest := #MAX_DATA_BUFFER - #statSend.tsendFct.dataOffset - 20;
                                   ELSE
                                       #statSend.tsendFct.dataLengthRest := #MAX_DATA_BUFFER - #statSend.tsendFct.dataOffset - 12;
                                   END_IF;

                                   //Calculate rest data from the total LCom message
                                   #tempUDint := #statSend.dataTelegram.totalMessageLength - #statSend.dataTelegram.messageOffset;

                                   //Calculate max. actual package length
                                   IF (#statSend.tsendFct.dataLengthRest > #diagnostics.partnerConfig.sizeOfReceiveBuffer) THEN
                                       #statMaxActPacketLength := #diagnostics.partnerConfig.sizeOfReceiveBuffer;
                                   ELSE
                                       #statMaxActPacketLength := #statSend.tsendFct.dataLengthRest;
                                   END_IF;

                                   //Rest data from the total LCom message, is greater than max. actual package length
                                   IF (#tempUDint > #statMaxActPacketLength) THEN
                                       #statSend.dataTelegram.actPackageLength := #statMaxActPacketLength;
                                   ELSE
                                       #statSend.dataTelegram.actPackageLength := #tempUDint;
                                   END_IF;

                                   #statSend.tsendFct.dataLengthRest := 0;
                                   //Build header from data telegram
                                   #statSend.tsendFct.data[#statSend.tsendFct.dataOffset] := #statSend.dataTelegram.LComVersion;
                                   #statSend.tsendFct.data[#statSend.tsendFct.dataOffset + 1] := #statSend.dataTelegram.telegramType;
                                   #statSend.tsendFct.data[#statSend.tsendFct.dataOffset + 2] := #statSend.dataTelegram.messageCounter;
                                   #statSend.tsendFct.data[#statSend.tsendFct.dataOffset + 3] := #statSend.dataTelegram.ackMessageCounter;

                                   #statSend.tsendFct.data[#statSend.tsendFct.dataOffset + 4] := #statSend.dataTelegram.messageOffset.%B3;
                                   #statSend.tsendFct.data[#statSend.tsendFct.dataOffset + 5] := #statSend.dataTelegram.messageOffset.%B2;
                                   #statSend.tsendFct.data[#statSend.tsendFct.dataOffset + 6] := #statSend.dataTelegram.messageOffset.%B1;
                                   #statSend.tsendFct.data[#statSend.tsendFct.dataOffset + 7] := #statSend.dataTelegram.messageOffset.%B0;

                                   #statSend.tsendFct.data[#statSend.tsendFct.dataOffset + 8] := #statSend.dataTelegram.ackMessageOffset.%B3;
                                   #statSend.tsendFct.data[#statSend.tsendFct.dataOffset + 9] := #statSend.dataTelegram.ackMessageOffset.%B2;
                                   #statSend.tsendFct.data[#statSend.tsendFct.dataOffset + 10] := #statSend.dataTelegram.ackMessageOffset.%B1;
                                   #statSend.tsendFct.data[#statSend.tsendFct.dataOffset + 11] := #statSend.dataTelegram.ackMessageOffset.%B0;

                                   #statSend.tsendFct.data[#statSend.tsendFct.dataOffset + 12] := #statSend.dataTelegram.actPackageLength.%B3;
                                   #statSend.tsendFct.data[#statSend.tsendFct.dataOffset + 13] := #statSend.dataTelegram.actPackageLength.%B2;
                                   #statSend.tsendFct.data[#statSend.tsendFct.dataOffset + 14] := #statSend.dataTelegram.actPackageLength.%B1;
                                   #statSend.tsendFct.data[#statSend.tsendFct.dataOffset + 15] := #statSend.dataTelegram.actPackageLength.%B0;

                                   #statSend.tsendFct.data[#statSend.tsendFct.dataOffset + 16] := #statSend.dataTelegram.totalMessageLength.%B3;
                                   #statSend.tsendFct.data[#statSend.tsendFct.dataOffset + 17] := #statSend.dataTelegram.totalMessageLength.%B2;
                                   #statSend.tsendFct.data[#statSend.tsendFct.dataOffset + 18] := #statSend.dataTelegram.totalMessageLength.%B1;
                                   #statSend.tsendFct.data[#statSend.tsendFct.dataOffset + 19] := #statSend.dataTelegram.totalMessageLength.%B0;

                                   //LCom V2
                                   IF (#diagnostics.statistics.activeLComVersion = #HEADER_V2) THEN
                                       //Calculate offset in the tcp send buffer
                                       #statSend.tsendFct.dataOffset := #statSend.tsendFct.dataOffset + 20;
                                   ELSE
                                       //LCom V1
                                       //MessageOffset
                                       #statSend.tsendFct.data[#statSend.tsendFct.dataOffset + 4] := #statSend.dataTelegram.messageOffset.%B1;
                                       #statSend.tsendFct.data[#statSend.tsendFct.dataOffset + 5] := #statSend.dataTelegram.messageOffset.%B0;
                                       //AckMessageOffset
                                       #statSend.tsendFct.data[#statSend.tsendFct.dataOffset + 6] := #statSend.dataTelegram.ackMessageOffset.%B1;
                                       #statSend.tsendFct.data[#statSend.tsendFct.dataOffset + 7] := #statSend.dataTelegram.ackMessageOffset.%B0;
                                       //ActPackageLength
                                       #statSend.tsendFct.data[#statSend.tsendFct.dataOffset + 8] := #statSend.dataTelegram.actPackageLength.%B1;
                                       #statSend.tsendFct.data[#statSend.tsendFct.dataOffset + 9] := #statSend.dataTelegram.actPackageLength.%B0;
                                       //TotalMessageLength
                                       #statSend.tsendFct.data[#statSend.tsendFct.dataOffset + 10] := #statSend.dataTelegram.totalMessageLength.%B1;
                                       #statSend.tsendFct.data[#statSend.tsendFct.dataOffset + 11] := #statSend.dataTelegram.totalMessageLength.%B0;
                                       //Calculate offset in the tcp send buffer
                                       #statSend.tsendFct.dataOffset := #statSend.tsendFct.dataOffset + 12;
                                   END_IF;

                                   //Store expected acknowledge message offset and time
                                   #statSend.expectedAck.package1.offset := #statSend.dataTelegram.messageOffset + #statSend.dataTelegram.actPackageLength;
                                   //Start expe. message Timer 1
                                   #instExpectedAckPackage1(IN := TRUE,
                                                            PT := #diagnostics.localConfig.sender.ackTimeout);

                                   #statSend.numberOfLComPackage := #statSend.numberOfLComPackage + 1;

                                   //Copy data from FB.sendBuffer
                                   #statRet := MOVE_BLK_VARIANT(SRC := #sendBuffer, COUNT := #statSend.dataTelegram.actPackageLength, SRC_INDEX := UDINT_TO_DINT(#statSend.userData.offset), DEST_INDEX := #statSend.tsendFct.dataOffset, DEST => #statSend.tsendFct.data);
                                   //Calculate offset in FB.sendBuffer
                                   #statSend.userData.offset := #statSend.userData.offset + #statSend.dataTelegram.actPackageLength;
                                   //Copy offset in telegram
                                   #statSend.dataTelegram.messageOffset := #statSend.userData.offset;
                                   //Calculate offset in the tcp send buffer
                                   #statSend.tsendFct.dataOffset := #statSend.tsendFct.dataOffset + UDINT_TO_UINT(#statSend.dataTelegram.actPackageLength);

                                   //All sent data is copied ?
                                   IF (#statSend.userData.offset = #statSend.dataTelegram.totalMessageLength) THEN
                                       //Yes
                                       #statState.comSender := #SEND_NO_DATA;
                                   ELSE
                                       ;//No --> Not all sent data has been copied
                                   END_IF;
                               ELSIF (#statState.comSender = #CYCLE
                                   AND
                                   (NOT #diagnostics.localConfig.connection.useLComProtocol)) THEN
                                   //---------------------------------------------------------------------
                                   //Send telegram without LCom protocol
                                   //---------------------------------------------------------------------
                                   #statState.sender := #SEND_DATA;

                                   //Calculate rest data from the total message
                                   IF ((#statSend.dataTelegram.totalMessageLength - #statSend.userData.offset) > #MAX_DATA_BUFFER) THEN
                                       #statSend.tsendFct.dataOffset := #MAX_DATA_BUFFER;
                                   ELSE
                                       #statSend.tsendFct.dataOffset := UDINT_TO_UINT(#statSend.dataTelegram.totalMessageLength - #statSend.userData.offset);
                                   END_IF;

                                   //Copy data from FB.sendBuffer
                                   #statRet := MOVE_BLK_VARIANT(SRC := #sendBuffer, COUNT := #statSend.tsendFct.dataOffset, SRC_INDEX := UDINT_TO_DINT(#statSend.userData.offset), DEST_INDEX := 0, DEST => #statSend.tsendFct.data);
                                   //Calculate offset in tcp send buffer
                                   #statSend.userData.offset := #statSend.userData.offset + #statSend.tsendFct.dataOffset;
                                   //End: Send telegram without LCom protocol
                               ELSE
                                   ;//Not in sending process 
                               END_IF;//End: Send telegram
                           END_REGION SEND_DATA_TELEGRAM

                       END_IF;//End: Connected
                   END_REGION HANDLE_SENDING

                   REGION SENDER_STATE_MACHINE
                       //---------------------------------------------------------------------
                       //State machine sender configuration
                       //---------------------------------------------------------------------
                       CASE #statState.cfgSender OF

                           #OPERATION:
                               ;//Sender configuration successful exchange
                           #STATE_WAIT:
                               ;
                           #STATE_INIT:

                               #statCompare.sender.cycleTime := #configuration.sender.cycleTime;
                               #statCompare.sender.ackTimeOut := #configuration.sender.ackTimeout;

                               //LCom Version V1.0
                               IF (#statActualLocalLComVersion = #HEADER_V1) THEN

                                   //Check max. cycleTime
                                   IF (#configuration.sender.cycleTime > T#65535ms) THEN

                                       #statDiag.bufferIndex := #statDiag.bufferIndex + 1;
                                       #statDiag.buffer[#statDiag.bufferIndex].additionalValue4 := #configuration.sender.cycleTime;
                                       #statSend.configTelegramV1.cycleTime := 65535;

                                       #statDiag.buffer[#statDiag.bufferIndex].status := #WARN_SEND_CYCLE_LIMITATION;
                                       #statDiag.buffer[#statDiag.bufferIndex].subFunctionErrorID := 16#0000;
                                       #statDiag.buffer[#statDiag.bufferIndex].additionalValue1 := 65535.0;
                                       #statDiag.buffer[#statDiag.bufferIndex].additionalValue2 := 0.0;
                                       #statDiag.buffer[#statDiag.bufferIndex].additionalValue3 := 0.0;
                                   ELSE
                                       #statSend.configTelegramV1.cycleTime := TIME_TO_UINT(#configuration.sender.cycleTime);
                                   END_IF;

                                   //Check max. ackTimeOut
                                   IF (#configuration.sender.ackTimeout > T#65535ms) THEN

                                       #statDiag.bufferIndex := #statDiag.bufferIndex + 1;
                                       #statDiag.buffer[#statDiag.bufferIndex].additionalValue4 := #configuration.sender.ackTimeout;
                                       #statSend.configTelegramV1.ackTimeOut := 65535;

                                       #statDiag.buffer[#statDiag.bufferIndex].status := #WARN_ACK_TIMEOUT_LIMITATION;
                                       #statDiag.buffer[#statDiag.bufferIndex].subFunctionErrorID := 16#0000;
                                       #statDiag.buffer[#statDiag.bufferIndex].additionalValue1 := 65535.0;
                                       #statDiag.buffer[#statDiag.bufferIndex].additionalValue2 := 0.0;
                                       #statDiag.buffer[#statDiag.bufferIndex].additionalValue3 := 0.0;
                                   ELSE
                                       #statSend.configTelegramV1.ackTimeOut := TIME_TO_UINT(#configuration.sender.ackTimeout);
                                   END_IF;
                               ELSE //LCom Version V2.0
                                   #statSend.configTelegramV2.cycleTime := #configuration.sender.cycleTime;
                                   #statSend.configTelegramV2.ackTimeOut := #configuration.sender.ackTimeout;
                               END_IF;

                               #statState.cfgSender := #SEND_CONFIG;

                           #SEND_CONFIG:
                               REGION SEND_CONFIG_TELEGRAM
                                   #statState.cfgSender := #STATE_WAIT;

                                   //LCom Version V1.0
                                   IF (#statActualLocalLComVersion = #HEADER_V1) THEN
                                       #statSend.tsendFct.data[#statSend.tsendFct.dataOffset] := #statSend.configTelegramV1.LComVersion;
                                       #statSend.tsendFct.data[#statSend.tsendFct.dataOffset + 1] := 16#02;
                                       #statSend.tsendFct.data[#statSend.tsendFct.dataOffset + 2] := #statSend.configTelegramV1.comMode;//ComMode
                                       #statSend.tsendFct.data[#statSend.tsendFct.dataOffset + 3] := #statSend.configTelegramV1.slidingWindow;//SlidingWindow
                                       //cycleTime
                                       #statSend.tsendFct.data[#statSend.tsendFct.dataOffset + 4] := #statSend.configTelegramV1.cycleTime.%B1;
                                       #statSend.tsendFct.data[#statSend.tsendFct.dataOffset + 5] := #statSend.configTelegramV1.cycleTime.%B0;
                                       //ackTimeOut
                                       #statSend.tsendFct.data[#statSend.tsendFct.dataOffset + 6] := #statSend.configTelegramV1.ackTimeOut.%B1;
                                       #statSend.tsendFct.data[#statSend.tsendFct.dataOffset + 7] := #statSend.configTelegramV1.ackTimeOut.%B0;
                                       //lifeSignCycle
                                       #statSend.tsendFct.data[#statSend.tsendFct.dataOffset + 8] := #statSend.configTelegramV1.lifeSignCycle.%B1;
                                       #statSend.tsendFct.data[#statSend.tsendFct.dataOffset + 9] := #statSend.configTelegramV1.lifeSignCycle.%B0;
                                       //status
                                       #statSend.tsendFct.data[#statSend.tsendFct.dataOffset + 10] := #statSend.configTelegramV1.status;
                                       //sendModeSyncTime
                                       #statSend.tsendFct.data[#statSend.tsendFct.dataOffset + 11] := #statSend.configTelegramV1.sendModeSyncTime;
                                       //maxSendDataLength
                                       #statSend.tsendFct.data[#statSend.tsendFct.dataOffset + 12] := #statSend.configTelegramV1.maxSendDataLength.%B1;
                                       #statSend.tsendFct.data[#statSend.tsendFct.dataOffset + 13] := #statSend.configTelegramV1.maxSendDataLength.%B0;
                                       //maxReceiveDataLength
                                       #statSend.tsendFct.data[#statSend.tsendFct.dataOffset + 14] := #statSend.configTelegramV1.maxReceiveDataLength.%B1;
                                       #statSend.tsendFct.data[#statSend.tsendFct.dataOffset + 15] := #statSend.configTelegramV1.maxReceiveDataLength.%B0;

                                       #statSend.tsendFct.data[#statSend.tsendFct.dataOffset + 16] := #statSend.configTelegramV1.LComVersion;
                                       #statSend.tsendFct.data[#statSend.tsendFct.dataOffset + 17] := 16#02;
                                       #statSend.tsendFct.data[#statSend.tsendFct.dataOffset + 18] := #statSend.configTelegramV1.comMode;//ComMode
                                       #statSend.tsendFct.data[#statSend.tsendFct.dataOffset + 19] := #statSend.configTelegramV1.slidingWindow;//SlidingWindow
                                       //cycleTime
                                       #statSend.tsendFct.data[#statSend.tsendFct.dataOffset + 20] := #statSend.configTelegramV1.cycleTime.%B1;
                                       #statSend.tsendFct.data[#statSend.tsendFct.dataOffset + 21] := #statSend.configTelegramV1.cycleTime.%B0;
                                       //ackTimeOut
                                       #statSend.tsendFct.data[#statSend.tsendFct.dataOffset + 22] := #statSend.configTelegramV1.ackTimeOut.%B1;
                                       #statSend.tsendFct.data[#statSend.tsendFct.dataOffset + 23] := #statSend.configTelegramV1.ackTimeOut.%B0;
                                       //lifeSignCycle
                                       #statSend.tsendFct.data[#statSend.tsendFct.dataOffset + 24] := #statSend.configTelegramV1.lifeSignCycle.%B1;
                                       #statSend.tsendFct.data[#statSend.tsendFct.dataOffset + 25] := #statSend.configTelegramV1.lifeSignCycle.%B0;
                                       //status
                                       #statSend.tsendFct.data[#statSend.tsendFct.dataOffset + 26] := #statSend.configTelegramV1.status;
                                       //sendModeSyncTime
                                       #statSend.tsendFct.data[#statSend.tsendFct.dataOffset + 27] := #statSend.configTelegramV1.sendModeSyncTime;
                                       //maxSendDataLength
                                       #statSend.tsendFct.data[#statSend.tsendFct.dataOffset + 28] := #statSend.configTelegramV1.maxSendDataLength.%B1;
                                       #statSend.tsendFct.data[#statSend.tsendFct.dataOffset + 29] := #statSend.configTelegramV1.maxSendDataLength.%B0;
                                       //maxReceiveDataLength
                                       #statSend.tsendFct.data[#statSend.tsendFct.dataOffset + 30] := #statSend.configTelegramV1.maxReceiveDataLength.%B1;
                                       #statSend.tsendFct.data[#statSend.tsendFct.dataOffset + 31] := #statSend.configTelegramV1.maxReceiveDataLength.%B0;
                                       //calculate new offset
                                       #statSend.tsendFct.dataOffset := #statSend.tsendFct.dataOffset + 32;
                                       #statState.sender := #SEND_CONFIG;

                                       #diagnostics.localConfig.sender.cycleTime := UINT_TO_TIME(#statSend.configTelegramV1.cycleTime);
                                       #diagnostics.localConfig.sender.ackTimeout := UINT_TO_TIME(#statSend.configTelegramV1.ackTimeOut);
                                   ELSE
                                       //LCom Version V2.0
                                       #statSend.tsendFct.data[#statSend.tsendFct.dataOffset] := #statSend.configTelegramV2.LComVersion;
                                       #statSend.tsendFct.data[#statSend.tsendFct.dataOffset + 1] := 16#02;
                                       //status
                                       #statSend.tsendFct.data[#statSend.tsendFct.dataOffset + 2] := #statSend.configTelegramV2.status;
                                       //sendModeSyncTime
                                       #statSend.tsendFct.data[#statSend.tsendFct.dataOffset + 3] := #statSend.configTelegramV2.sendModeSyncTime;
                                       //lifeSignCycle
                                       #tempDWord := TIME_TO_DWORD(#statSend.configTelegramV2.lifeSignCycle);
                                       #statSend.tsendFct.data[#statSend.tsendFct.dataOffset + 4] := #tempDWord.%B3;
                                       #statSend.tsendFct.data[#statSend.tsendFct.dataOffset + 5] := #tempDWord.%B2;
                                       #statSend.tsendFct.data[#statSend.tsendFct.dataOffset + 6] := #tempDWord.%B1;
                                       #statSend.tsendFct.data[#statSend.tsendFct.dataOffset + 7] := #tempDWord.%B0;
                                       //cycleTime
                                       #tempDWord := TIME_TO_DWORD(#statSend.configTelegramV2.cycleTime);
                                       #statSend.tsendFct.data[#statSend.tsendFct.dataOffset + 8] := #tempDWord.%B3;
                                       #statSend.tsendFct.data[#statSend.tsendFct.dataOffset + 9] := #tempDWord.%B2;
                                       #statSend.tsendFct.data[#statSend.tsendFct.dataOffset + 10] := #tempDWord.%B1;
                                       #statSend.tsendFct.data[#statSend.tsendFct.dataOffset + 11] := #tempDWord.%B0;
                                       //ackTimeOut
                                       #tempDWord := TIME_TO_DWORD(#statSend.configTelegramV2.ackTimeOut);
                                       #statSend.tsendFct.data[#statSend.tsendFct.dataOffset + 12] := #tempDWord.%B3;
                                       #statSend.tsendFct.data[#statSend.tsendFct.dataOffset + 13] := #tempDWord.%B2;
                                       #statSend.tsendFct.data[#statSend.tsendFct.dataOffset + 14] := #tempDWord.%B1;
                                       #statSend.tsendFct.data[#statSend.tsendFct.dataOffset + 15] := #tempDWord.%B0;
                                       //maxSendDataLength
                                       #statSend.tsendFct.data[#statSend.tsendFct.dataOffset + 16] := #statSend.configTelegramV2.maxSendDataLength.%B3;
                                       #statSend.tsendFct.data[#statSend.tsendFct.dataOffset + 17] := #statSend.configTelegramV2.maxSendDataLength.%B2;
                                       #statSend.tsendFct.data[#statSend.tsendFct.dataOffset + 18] := #statSend.configTelegramV2.maxSendDataLength.%B1;
                                       #statSend.tsendFct.data[#statSend.tsendFct.dataOffset + 19] := #statSend.configTelegramV2.maxSendDataLength.%B0;
                                       //maxReceiveDataLength
                                       #statSend.tsendFct.data[#statSend.tsendFct.dataOffset + 20] := #statSend.configTelegramV2.maxReceiveDataLength.%B3;
                                       #statSend.tsendFct.data[#statSend.tsendFct.dataOffset + 21] := #statSend.configTelegramV2.maxReceiveDataLength.%B2;
                                       #statSend.tsendFct.data[#statSend.tsendFct.dataOffset + 22] := #statSend.configTelegramV2.maxReceiveDataLength.%B1;
                                       #statSend.tsendFct.data[#statSend.tsendFct.dataOffset + 23] := #statSend.configTelegramV2.maxReceiveDataLength.%B0;

                                       //calculate new offset
                                       #statSend.tsendFct.dataOffset := #statSend.tsendFct.dataOffset + 24;
                                       #statState.sender := #SEND_CONFIG;

                                       #diagnostics.localConfig.sender.cycleTime := #statSend.configTelegramV2.cycleTime;
                                       #diagnostics.localConfig.sender.ackTimeout := #statSend.configTelegramV2.ackTimeOut;

                                       IF #diagnostics.statistics.activeLComVersion = #HEADER_V2 THEN
                                           #connected := #statConnected := TRUE;
                                           #diagnostics.statistics.LComProtocolUsed := TRUE;
                                           #diagnostics.statistics.activeLComVersion := #HEADER_V2;
                                           #statState.cfgSender := #OPERATION;

                                           //Write diagnostics
                                           #statDiag.bufferIndex := #statDiag.bufferIndex + 1;
                                           #statDiag.buffer[#statDiag.bufferIndex].status := #STATUS_CONNECTED_V2;
                                           #statDiag.buffer[#statDiag.bufferIndex].subFunctionErrorID := 16#0000;
                                           #statDiag.buffer[#statDiag.bufferIndex].additionalValue1 := 0.0;
                                           #statDiag.buffer[#statDiag.bufferIndex].additionalValue2 := 0.0;
                                           #statDiag.buffer[#statDiag.bufferIndex].additionalValue3 := 0.0;
                                           #statDiag.buffer[#statDiag.bufferIndex].additionalValue4 := T#0ms;
                                       END_IF;
                                   END_IF;

                                   #statCompare.sender.cycleTime := #configuration.sender.cycleTime;
                                   #statCompare.sender.ackTimeOut := #configuration.sender.ackTimeout;
                               END_REGION SEND_CONFIG_TELEGRAM

                           #ERROR_STATE:
                               ;
                           ELSE
                               ;// Statement section ELSE
                       END_CASE;
                   END_REGION SENDER_STATE_MACHINE

                   REGION SEND_LIFESIGN
                       //No telegram 1,2,5 or 10 to  be sent, therefore check whether life sign tel. must be sent
                       IF (#statState.sender = #STATE_INACTIVE
                           AND
                           (#diagnostics.localConfig.connection.lifeSignCycleTime <> T#0ms)
                           AND
                           #diagnostics.localConfig.connection.useLComProtocol)
                       THEN
                           #instLocalLifeSignCycleTimer(IN := TRUE,
                                                        PT := #diagnostics.localConfig.connection.lifeSignCycleTime);

                           IF (#instLocalLifeSignCycleTimer.Q)
                           THEN

                               //LCom Version V1.0
                               IF (#statActualLocalLComVersion = #HEADER_V1) THEN

